Fanuc KAREL source: KT00896.KL

PROGRAM KT00896
%NOLOCKGROUP
VAR
  P1: JOINTPOS
  P2: JOINTPOS
  OUT: BOOLEAN
BEGIN
  OUT = IN_RANGE(P1)
END KT00896
